(* IEC 61131-3 sources: daoli-st-library/DL_Process (part 4) *)

(* ---- FB_DL_MultiTankBlendSeq.st ---- *)
(*
  ============================================================
  组件名 : FB_DL_MultiTankBlendSeq
  分类   : DL_Process
  功能   : 多罐调和批次序列（A 进料 → B 进料 → 循环调和 → 取样 → 排料 → 完成），含超容、进料超时、收敛超时、取样超时、排料超时、人工中止、配方无效共七类故障锁存
  开源溯源 : internal-design（本轮无外部代码逐行引用）；参考语义 : 无外部参考
  复杂度 : C4
  版本   : 1.0.0
  ============================================================
*)

(*-----------------------------------------------------------------------------
 * 状态迁移表（ENUM 成员 → 出口；每成员均有可到达出口，零无界驻留相）：
 *   eIdle      → eFillA  : bStart 且 bRecipeValid 且组态闸通过 且 总量 ≤ rMaxVolume
 *   eIdle      ── 保持，直到 bStart（待机相以启动命令为唯一出口，属许可型驻留）
 *   eFillA     → eFillB  : rVolAct ≥ rVolA_sp（含 1E-6 容差）
 *   eFillA     → eFault  : tonFill.Q（码 1）｜bAbort 沿（码 5）｜rVolAct > rMaxVolume（码 4）｜bStart 撤除（无码回空闲）
 *   eFillB     → eCirculate : rVolAct ≥ (rVolA_sp + rVolB_sp) - 1E-6
 *   eFillB     → eFault  : tonFill.Q（码 1）｜bAbort 沿（码 5）｜超容（码 4）｜组态闸失效（码 6）
 *   eCirculate → eSample : 温度与浓度同时进带并持续 tCircStable（tonStable.Q）
 *   eCirculate → eFault  : tonCirc.Q（码 2）｜bAbort 沿（码 5）
 *   eSample    → eRelease : bSampleDone（外部取样完成电平）
 *   eSample    → eFault   : tonSample.Q（码 3）｜bAbort 沿（码 5）
 *   eRelease   → eDone    : bLevelLow（低液位信号，排料到位）
 *   eRelease   → eFault   : tonRelease.Q（码 7）｜bAbort 沿（码 5）
 *   eDone      → eIdle    : bStart 撤除（完成相以撤令为唯一出口，属人工确认型驻留）
 *   eFault     → eIdle    : bAbort 上升沿 或（bStart = FALSE 且 bAbort = FALSE）
 *   ELSE（非法枚举值，非任何成员）→ eFault（码 8）
 *
 * 故障码表（nFaultCode，0 = 无故障；非首码均附「现有输出不可观测」反证句，R90）：
 *   1 进料超时      : tFillTimeout 覆盖 eFillA + eFillB（进 eFillA 时计时器自然复位）。
 *   2 循环收敛超时  : 反证——eFault 相动作全撤后 bValveA/bValveB/bAgitator/bDischarge 全 FALSE、
 *                     eState 同为 eFault，复用码 1 会使「调和未收敛」与「进料过慢」在 HMI 上不可区分。
 *   3 取样超时      : 反证——取样相外部回执缺失，阀位与搅拌状态在故障撤除后与码 2 完全同形，
 *                     复用码 2 会把「外部取样单元不回报」误判为工艺收敛失败，运维方向相悖。
 *   4 超罐容        : 反证——超容判据在进料前即可成立（无阀位动作、无累计体积），
 *                     复用码 1 会把「配方总量超罐容」报成「进料慢」，掩盖配方错误。
 *   5 人工中止      : 反证——操作员主动撤令属安全审计事件，与任何超时码的因果主体不同，
 *                     合并后无法区分「设备不动」与「人按了停」。
 *   6 配方无效      : 反证——非法配方在进料前拦截，此时无累计体积、无阀位输出，
 *                     与超时类码位的时序签名互斥，必须独立成码以便前置拦截可被观测。
 *   7 排料超时      : 反证——排料相 bDischarge 独占且 bLevelLow 缺失，故障撤除后与码 1/2/3 的
 *                     观测量全同，复用码 1 会让运维去查进料阀而非排料阀。
 *   8 非法状态枚举  : 反证——非法枚举值为程序缺陷而非工艺事件，必须与现场工艺故障分离，
 *                     否则固件错误会被误排为设备故障。
 *
 * 依赖     : 仅 IEC 61131-3 标准库（TON / R_TRIG / ABS / LIMIT），零厂商私有库
 * 分工声明 : 循环泵输出不在本件接口（上层以 eState = eCirculate 派生泵命令）；
 *            温度/浓度闭环调节归温控件与浓度调节件；本件只做批次时序与保护，不做连续调节。
 * 归属     : E_DL_BlendState 归属本文件（全库唯一定义，R264；引用件只引用不重声明）。
 * 修订历史 : 2026-11-25  v1.0.0  首版（编码席 dlf-plc-coder，第二批 C4）
 *----------------------------------------------------------------------------*)

(*-----------------------------------------------------------------------------
 * 边界与红线自检：
 * ① 六个 TON 与一个 R_TRIG 全部在 CASE 外无条件周期调用（R7）；时间类 IN 均含 NOT .Q 自复位项
 *    与 NOT 故障锁存项（R188 / FB50-1③），CASE 内只读 .Q。
 * ② 出口命令（bValveA/bValveB/bAgitator/bDischarge/bSampleReq）在段 0 每拍预置 FALSE，
 *    CASE 内只置 TRUE —— eIdle 与 eFault 相零残留（上轮 MAJOR「故障后残留旧输出」型缺陷已封堵）。
 * ③ bDone 由相位派生（bDone := _eState = eDone），不是单拍脉冲，从结构上排除「同拍置位又撤销」（FB33-1）。
 * ④ 故障码 _nFault 一律锁存至 eFault 复位分支，故障相内不按当下输入重算（FB33-1③ / R152）。
 * ⑤ 除零防护：进度式除子 _rVolTotal 先过 > 1E-6 与 _bCfgOk 双检（R4）。
 * ⑥ 相内等待出口 ≥2（R98）：eSample = bSampleDone ｜ tonSample.Q ｜ bAbort 沿 ｜ bStart 撤除；
 *    eRelease = bLevelLow ｜ tonRelease.Q ｜ bAbort 沿 ｜ bStart 撤除。
 * ⑦ 组态域闸：参与任何判据换算的 10 个浮点入参全部显式枚举（含 rMaxVolume），NaN 用自反比较、
 *    Inf 用差值自减双判（R151 / R79），非有限不入保持槽。
 * ⑧ 零全局耦合：无 GVL / VAR_EXTERNAL / %I / %Q（R1 / R2）。
 * ⑨ 相位写入点共三处且互斥：段 3（bAbort 沿只置锁存，不写相位）、段 4 CASE、段 6 迁移闸。
 *----------------------------------------------------------------------------*)

TYPE E_DL_BlendState :
(
    eIdle      := 0, // 空闲：全部阀位关闭，等启动与配方有效 idle: all valves closed, waiting for start and a valid recipe
    eFillA     := 1, // A 罐进料相：开 A 阀累计至 rVolA_sp fill A: A valve open until rVolA_sp is reached
    eFillB     := 2, // B 罐进料相：开 B 阀累计至 A+B 总量 fill B: B valve open until the A+B total is reached
    eCirculate := 3, // 循环调和相：搅拌运行，温度与浓度双判进带 circulate: agitation with temperature and concentration both inside band
    eSample    := 4, // 取样相：置取样请求等外部完成 sample: sample request raised, waiting for the external completion
    eRelease   := 5, // 排料相：开排料阀至低液位 release: discharge valve open until the low level signal
    eFault     := 6, // 故障锁存相：全部阀位撤除，只由复位出口迁出 fault: all valves withdrawn, left only by the reset outlet
    eDone      := 7  // 批次完成相：bStart 撤除后回空闲 done: returns to idle when bStart is withdrawn
);
END_TYPE

FUNCTION_BLOCK FB_DL_MultiTankBlendSeq
VAR_INPUT
    bStart          : BOOL := FALSE;          // 启动/运行许可（电平）：撤除即安全停机回空闲 [bool] start and run permissive, a dropped level stops safely
    bAbort          : BOOL := FALSE;          // 人工中止（上升沿）：置故障码 5 并锁存 [bool] manual abort rising edge, latches fault code 5
    bRecipeValid    : BOOL := FALSE;          // 配方有效回执：FALSE 时禁止启动并置码 6 [bool] recipe valid receipt, FALSE blocks the start with code 6
    rVolA_sp        : REAL := 0.0;            // A 组分配方体积设定 [m3] recipe volume setpoint of component A [m3]
    rVolB_sp        : REAL := 0.0;            // B 组分配方体积设定 [m3] recipe volume setpoint of component B [m3]
    rVolAct         : REAL := 0.0;            // 当前累计进料量（A+B 合计）[m3] accumulated feed volume of A plus B [m3]
    rTempAct        : REAL := 0.0;            // 混合物实测温度 [degC] measured blend temperature [degC]
    rTempSp         : REAL := 0.0;            // 调和温度设定 [degC] blend temperature setpoint [degC]
    rTempBand       : REAL := 0.0;            // 温度进带允许偏差，域 > 1E-6 [K] temperature band tolerance, domain > 1E-6 [K]
    rConcAct        : REAL := 0.0;            // 混合物实测浓度 [%] measured blend concentration [%]
    rConcSp         : REAL := 0.0;            // 调和浓度设定 [%] blend concentration setpoint [%]
    rConcBand       : REAL := 0.0;            // 浓度进带允许偏差，域 > 1E-6 [%] concentration band tolerance, domain > 1E-6 [%]
    tFillTimeout    : TIME := T#10M;          // 进料总超时窗，覆盖 eFillA + eFillB [s] total feed timeout covering fill A and fill B [s]
    tCircTimeout    : TIME := T#30M;          // 循环调和相超时窗 [s] circulation phase timeout window [s]
    tSampleTimeout  : TIME := T#5M;           // 取样相等待外部回执超时窗 [s] sample phase external receipt timeout [s]
    rMaxVolume      : REAL := 10.0;           // 罐体最大有效容积，域 > 0 [m3] tank maximum usable volume, domain > 0 [m3]
    bSampleDone     : BOOL := FALSE;          // 外部取样完成回执（电平）[bool] external sampling done receipt level
    bLevelLow       : BOOL := FALSE;          // 排料低液位信号（排料到位）[bool] discharge low level signal
    tCircStable     : TIME := T#15S;          // 温度与浓度同时在带内的持续确认窗 [s] continuous in-band confirmation window [s]
    tReleaseTimeout : TIME := T#15M;          // 排料相超时窗（低液位不到的兜底）[s] release phase timeout fallback [s]
END_VAR
VAR_OUTPUT
    bValveA      : BOOL;                      // A 组分进料阀命令（段 0 预置，CASE 只置位）[bool] component A feed valve command
    bValveB      : BOOL;                      // B 组分进料阀命令（段 0 预置，CASE 只置位）[bool] component B feed valve command
    bAgitator    : BOOL;                      // 搅拌器命令（循环相与取样相保持开）[bool] agitator command, held in circulation and sampling
    bDischarge   : BOOL;                      // 排料阀命令（仅排料相）[bool] discharge valve command, release phase only
    bSampleReq   : BOOL;                      // 取样请求（仅取样相，电平保持）[bool] sample request, level held in the sample phase
    eState       : E_DL_BlendState;           // 相位出口（段 7 单点映射）[-] phase outlet mapped once in section 7
    bDone        : BOOL;                      // 批次完成（由相位派生，非单拍脉冲）[bool] batch done, derived from the phase as a level
    nFaultCode   : INT;                       // 故障码 0 无 1 进料超时 2 收敛超时 3 取样超时 4 超容 5 人工中止 6 配方无效 7 排料超时 8 非法状态 [码] fault code
    rProgressPct : REAL;                      // 进料完成度 0..100（其后各相恒 100）[%] feed completion percentage, constant 100 in later phases [%]
    bError       : BOOL;                      // 故障锁存标志（取锁存位，R45 配对出口）[bool] fault latch flag used as the paired outlet
END_VAR
VAR
    _eState       : E_DL_BlendState := E_DL_BlendState.eIdle;   // 内部相位（CASE 唯一比较目标）[-] internal phase compared by the CASE
    _bFaultLatch  : BOOL := FALSE;                              // 故障锁存位（仅复位出口清除）[bool] fault latch, cleared only by the reset outlet
    _nFault       : INT := 0;                                   // 锁存故障码（故障期回放，不按当下输入重算）[码] latched fault code replayed during the fault phase
    _bCfgOk       : BOOL := FALSE;                              // 组态与入参域闸通过标志 [bool] configuration and input domain gate flag
    _bRunActive   : BOOL := FALSE;                              // 运行相关相标志（进料到排料）[bool] running phase flag from fill to release
    _bInBand      : BOOL := FALSE;                               // 温度与浓度同时进带标志 [bool] both temperature and concentration inside band
    _bValveA      : BOOL := FALSE;                              // 内部 A 阀命令状态 [bool] internal A valve command state
    _bValveB      : BOOL := FALSE;                              // 内部 B 阀命令状态 [bool] internal B valve command state
    _bAgitator    : BOOL := FALSE;                              // 内部搅拌命令状态 [bool] internal agitator command state
    _bDischarge   : BOOL := FALSE;                              // 内部排料阀命令状态 [bool] internal discharge valve command state
    _bSampleReq   : BOOL := FALSE;                              // 内部取样请求状态 [bool] internal sample request state
    _rVolTotal    : REAL := 0.0;                                // 配方总量 = A + B [m3] recipe total volume of A plus B [m3]
    _rProg        : REAL := 0.0;                                // 进料完成度中间量 [%] feed completion intermediate value [%]
    rtAbort       : R_TRIG;                                     // bAbort 上升沿实例（段 2 无条件调用）[bool] abort rising edge instance
    tonFill       : TON;                                        // 进料总超时计时（覆盖两进料相，段 2 无条件调用）[s] total feed timeout covering both fill phases
    tonCirc       : TON;                                        // 循环调和相超时计时（段 2 无条件调用）[s] circulation timeout
    tonStable     : TON;                                        // 双判进带持续确认计时（段 2 无条件调用）[s] in-band persistence timer
    tonSample     : TON;                                        // 取样相等待回执超时计时（段 2 无条件调用）[s] sample receipt timeout
    tonRelease    : TON;                                        // 排料相超时计时（段 2 无条件调用）[s] release timeout
END_VAR
VAR CONSTANT
    DL_BLD_ZERO     : REAL := 0.0;        // 浮点零基准 [m3] float zero base
    DL_BLD_ONE      : REAL := 1.0;        // 浮点一基准 [%] float one base
    DL_BLD_HUNDRED  : REAL := 100.0;      // 百分比满量程 [%] percent full scale
    DL_BLD_EPS      : REAL := 1.0E-6;     // 体积与宽容差基准 [m3] volume and band tolerance base
    DL_BLD_T_MIN    : TIME := T#100MS;    // 时间参数下限 [s] lower bound of the time parameters
    DL_BLD_T_MAX    : TIME := T#4H;       // 时间参数上限 [s] upper bound of the time parameters
END_VAR

(* —— 段 0：出口命令预置与派生量计算（CASE 内只置 TRUE，杜绝故障相残留） —— *)
_bValveA    := FALSE;                                               // A 阀命令每拍先撤 [bool] A valve withdrawn first each scan
_bValveB    := FALSE;                                               // B 阀命令每拍先撤 [bool] B valve withdrawn first each scan
_bAgitator  := FALSE;                                               // 搅拌命令每拍先撤 [bool] agitator withdrawn first each scan
_bDischarge := FALSE;                                               // 排料阀命令每拍先撤 [bool] discharge withdrawn first each scan
_bSampleReq := FALSE;                                               // 取样请求每拍先撤 [bool] sample request withdrawn first each scan
_rProg      := DL_BLD_ZERO;                                         // 进度中间量每拍清零 [%] progress intermediate cleared each scan
_rVolTotal  := rVolA_sp + rVolB_sp;                                 // 配方总量求和 [m3] recipe total volume
_bRunActive := (_eState = E_DL_BlendState.eFillA) OR (_eState = E_DL_BlendState.eFillB)
               OR (_eState = E_DL_BlendState.eCirculate) OR (_eState = E_DL_BlendState.eSample)
               OR (_eState = E_DL_BlendState.eRelease);             // 运行相关相标志（用状态量，R99）[bool] running phase flag from the state
_bInBand    := FALSE;                                               // 进带标志复位 [bool] in-band flag reset
IF (rTempBand > DL_BLD_ZERO) AND (rConcBand > DL_BLD_ZERO) THEN
    IF (ABS(rTempAct - rTempSp) <= rTempBand) AND (ABS(rConcAct - rConcSp) <= rConcBand) THEN
        _bInBand := TRUE;                                           // 双判同时进带 [bool] both criteria inside band
    END_IF
END_IF

(* —— 段 1：组态域闸与容量保护（十个浮点入参全枚举，非有限双判 R151 / R79） —— *)
_bCfgOk := TRUE;                                                    // 组态闸标志初值 [bool] configuration flag initial value
IF (rVolA_sp <> rVolA_sp) OR ((rVolA_sp - rVolA_sp) <> DL_BLD_ZERO)
   OR (rVolB_sp <> rVolB_sp) OR ((rVolB_sp - rVolB_sp) <> DL_BLD_ZERO)
   OR (rVolAct <> rVolAct) OR ((rVolAct - rVolAct) <> DL_BLD_ZERO)
   OR (rMaxVolume <> rMaxVolume) OR ((rMaxVolume - rMaxVolume) <> DL_BLD_ZERO)
   OR (rTempAct <> rTempAct) OR ((rTempAct - rTempAct) <> DL_BLD_ZERO)
   OR (rTempSp <> rTempSp) OR ((rTempSp - rTempSp) <> DL_BLD_ZERO)
   OR (rTempBand <> rTempBand) OR ((rTempBand - rTempBand) <> DL_BLD_ZERO)
   OR (rConcAct <> rConcAct) OR ((rConcAct - rConcAct) <> DL_BLD_ZERO)
   OR (rConcSp <> rConcSp) OR ((rConcSp - rConcSp) <> DL_BLD_ZERO)
   OR (rConcBand <> rConcBand) OR ((rConcBand - rConcBand) <> DL_BLD_ZERO) THEN
    _bCfgOk := FALSE;                                               // 非有限入参：拒收（NaN 自反 + Inf 差值自减）[bool] non finite input rejected
END_IF
IF _bCfgOk THEN
    IF (rVolA_sp < DL_BLD_ZERO) OR (rVolB_sp < DL_BLD_ZERO) OR (rMaxVolume <= DL_BLD_ZERO) THEN
        _bCfgOk := FALSE;                                           // 负体积或非正罐容 [bool] negative volume or non positive capacity
    ELSIF (_rVolTotal <= DL_BLD_ZERO) THEN
        _bCfgOk := FALSE;                                           // 配方总量为零 [bool] zero recipe total volume
    ELSIF (rTempBand < DL_BLD_EPS) OR (rConcBand < DL_BLD_EPS) THEN
        _bCfgOk := FALSE;                                           // 容差带为零或负 [bool] zero or negative tolerance band
    ELSIF (tFillTimeout < DL_BLD_T_MIN) OR (tFillTimeout > DL_BLD_T_MAX) THEN
        _bCfgOk := FALSE;                                           // 进料超时越域 [bool] feed timeout out of domain
    ELSIF (tCircTimeout < DL_BLD_T_MIN) OR (tCircTimeout > DL_BLD_T_MAX) THEN
        _bCfgOk := FALSE;                                           // 循环超时越域 [bool] circulation timeout out of domain
    ELSIF (tSampleTimeout < DL_BLD_T_MIN) OR (tSampleTimeout > DL_BLD_T_MAX) THEN
        _bCfgOk := FALSE;                                           // 取样超时越域 [bool] sample timeout out of domain
    ELSIF (tCircStable < DL_BLD_T_MIN) OR (tCircStable > DL_BLD_T_MAX) THEN
        _bCfgOk := FALSE;                                           // 进带确认窗越域 [bool] in-band window out of domain
    ELSIF (tReleaseTimeout < DL_BLD_T_MIN) OR (tReleaseTimeout > DL_BLD_T_MAX) THEN
        _bCfgOk := FALSE;                                           // 排料超时越域 [bool] release timeout out of domain
    ELSIF NOT bRecipeValid THEN
        _bCfgOk := FALSE;                                           // 配方无效回执为假 [bool] recipe valid receipt is false
    END_IF
END_IF
IF (NOT _bCfgOk) AND (NOT _bFaultLatch) AND (bStart OR _bRunActive) THEN
    _nFault      := 6;                                              // 故障级：配方无效 / 参数非法 [码] fault: invalid recipe or parameter
    _bFaultLatch := TRUE;                                           // 置故障锁存 [bool] latch the fault
    bError       := TRUE;                                           // R45 配对：故障标志同拍置位 [bool] paired error flag
END_IF
IF (NOT _bFaultLatch) AND (bStart OR _bRunActive) THEN
    IF _rVolTotal > rMaxVolume THEN
        _nFault      := 4;                                          // 故障级：配方总量超罐容 [码] fault: recipe total exceeds tank volume
        _bFaultLatch := TRUE;                                       // 置故障锁存 [bool] latch the fault
        bError       := TRUE;                                       // R45 配对：故障标志同拍置位 [bool] paired error flag
    END_IF
END_IF

(* —— 段 2：边沿与定时器（CASE 外无条件周期调用，R7；IN 含 NOT .Q 自复位与 NOT 锁存，R188） —— *)
rtAbort(CLK := bAbort);                                             // bAbort 边沿无条件刷新 [bool] abort edge refreshed unconditionally
tonFill(IN := ((_eState = E_DL_BlendState.eFillA) OR (_eState = E_DL_BlendState.eFillB))
              AND (NOT tonFill.Q) AND (NOT _bFaultLatch),
        PT := tFillTimeout);                                        // 进料总超时（跨两相累计，进相自然复位）[s] total feed timeout across both phases
tonCirc(IN := (_eState = E_DL_BlendState.eCirculate) AND (NOT tonCirc.Q) AND (NOT _bFaultLatch),
        PT := tCircTimeout);                                        // 循环调和超时 [s] circulation timeout
tonStable(IN := (_eState = E_DL_BlendState.eCirculate) AND _bInBand AND (NOT tonStable.Q)
               AND (NOT _bFaultLatch),
          PT := tCircStable);                                       // 双判进带持续确认 [s] in-band persistence confirmation
tonSample(IN := (_eState = E_DL_BlendState.eSample) AND (NOT tonSample.Q) AND (NOT _bFaultLatch),
          PT := tSampleTimeout);                                    // 取样回执超时 [s] sample receipt timeout
tonRelease(IN := (_eState = E_DL_BlendState.eRelease) AND (NOT tonRelease.Q) AND (NOT _bFaultLatch),
           PT := tReleaseTimeout);                                  // 排料超时 [s] release timeout

(* —— 段 3：人工中止优先消化（置锁存不写相位，迁相由段 6 统一执行，R21 / R275） —— *)
IF rtAbort.Q AND (NOT _bFaultLatch) THEN
    _nFault      := 5;                                              // 故障级：人工中止 [码] fault: manual abort
    _bFaultLatch := TRUE;                                           // 置故障锁存 [bool] latch the fault
    bError       := TRUE;                                           // R45 配对：故障标志同拍置位 [bool] paired error flag
END_IF

(* —— 段 4：主状态机（相位写入点之二；每成员独立标签，ELSE 只兜非法值） —— *)
CASE _eState OF
E_DL_BlendState.eIdle :                                             // 空闲相：全部阀位已撤，等启动与配方许可
    IF bStart AND _bCfgOk AND (NOT bAbort) AND (NOT _bFaultLatch) THEN
        _eState := E_DL_BlendState.eFillA;                          // 迁移：进入 A 进料相（次拍开阀）[phase] move to fill A
    END_IF

E_DL_BlendState.eFillA :                                            // A 进料相：开 A 阀
    _bValveA := TRUE;                                               // 开 A 组分进料阀 [bool] open the component A feed valve
    IF rVolAct >= (rVolA_sp - DL_BLD_EPS) THEN
        _eState := E_DL_BlendState.eFillB;                          // 迁移：A 组分量已到位 [phase] component A volume reached
    ELSIF rVolAct > rMaxVolume THEN
        _nFault      := 4;                                          // 故障级：累计体积超罐容 [码] fault: accumulated volume over capacity
        _bFaultLatch := TRUE;                                       // 置故障锁存 [bool] latch the fault
        bError       := TRUE;                                       // R45 配对：故障标志同拍置位 [bool] paired error flag
    END_IF

E_DL_BlendState.eFillB :                                            // B 进料相：开 B 阀至总量
    _bValveB := TRUE;                                               // 开 B 组分进料阀 [bool] open the component B feed valve
    IF rVolAct >= (_rVolTotal - DL_BLD_EPS) THEN
        _eState := E_DL_BlendState.eCirculate;                      // 迁移：总量到位进入循环调和 [phase] total volume reached, start circulation
    ELSIF rVolAct > rMaxVolume THEN
        _nFault      := 4;                                          // 故障级：累计体积超罐容 [码] fault: accumulated volume over capacity
        _bFaultLatch := TRUE;                                       // 置故障锁存 [bool] latch the fault
        bError       := TRUE;                                       // R45 配对：故障标志同拍置位 [bool] paired error flag
    END_IF

E_DL_BlendState.eCirculate :                                        // 循环调和相：搅拌运行，温度与浓度双判
    _bAgitator := TRUE;                                             // 搅拌保持开（保证均质）[bool] agitator held on for homogeneity
    IF tonStable.Q THEN
        _eState := E_DL_BlendState.eSample;                         // 迁移：双判进带持续满足 [phase] both criteria held inside band
    END_IF

E_DL_BlendState.eSample :                                           // 取样相：请求外部取样并等待回执
    _bAgitator  := TRUE;                                            // 取样期间保持搅拌（样品代表性）[bool] agitator held during sampling
    _bSampleReq := TRUE;                                            // 置取样请求（电平保持）[bool] sample request level held
    IF bSampleDone THEN
        _eState := E_DL_BlendState.eRelease;                        // 迁移（出口 1）：外部取样完成 [phase] external sampling completed
    END_IF

E_DL_BlendState.eRelease :                                          // 排料相：开排料阀至低液位
    _bDischarge := TRUE;                                            // 开排料阀（搅拌停，避免抽空涡流）[bool] open the discharge valve
    IF bLevelLow THEN
        _eState := E_DL_BlendState.eDone;                           // 迁移（出口 1）：低液位到位 [phase] low level reached
    END_IF

E_DL_BlendState.eDone :                                             // 完成相：bDone 由相位派生，等撤令
    IF NOT bStart THEN
        _eState := E_DL_BlendState.eIdle;                           // 迁移：撤除启动命令回空闲 [phase] start withdrawn, back to idle
    END_IF

E_DL_BlendState.eFault :                                            // 故障锁存相：阀位已由段 6 全撤
    IF rtAbort.Q OR ((NOT bStart) AND (NOT bAbort)) THEN
        _bFaultLatch := FALSE;                                      // 复位出口：清故障锁存 [bool] clear the fault latch
        _nFault      := 0;                                          // 复位出口：清故障码 [码] clear the fault code
        _eState      := E_DL_BlendState.eIdle;                      // 复位出口：迁回空闲 [phase] back to idle
    END_IF

ELSE                                                                // 非法枚举值兜底（R6 / FB32-5）
    IF NOT _bFaultLatch THEN
        _nFault      := 8;                                          // 故障级：非法状态枚举值 [码] fault: illegal state enum value
        _bFaultLatch := TRUE;                                       // 置故障锁存 [bool] latch the fault
        bError       := TRUE;                                       // R45 配对：故障标志同拍置位 [bool] paired error flag
    END_IF
    _eState := E_DL_BlendState.eFault;                              // 非法值一律落安全相 [phase] illegal value falls into the safe phase
END_CASE

(* —— 段 5：超时看门狗锁存（本拍合法事件优先于超时：状态已迁出则该相看门狗不生效，R275） —— *)
IF tonFill.Q AND (NOT _bFaultLatch)
   AND ((_eState = E_DL_BlendState.eFillA) OR (_eState = E_DL_BlendState.eFillB)) THEN
    _nFault      := 1;                                              // 故障级：进料超时 [码] fault: feed timeout
    _bFaultLatch := TRUE;                                           // 置故障锁存 [bool] latch the fault
    bError       := TRUE;                                           // R45 配对：故障标志同拍置位 [bool] paired error flag
END_IF
IF tonCirc.Q AND (NOT _bFaultLatch) AND (_eState = E_DL_BlendState.eCirculate) THEN
    _nFault      := 2;                                              // 故障级：循环收敛超时 [码] fault: circulation convergence timeout
    _bFaultLatch := TRUE;                                           // 置故障锁存 [bool] latch the fault
    bError       := TRUE;                                           // R45 配对：故障标志同拍置位 [bool] paired error flag
END_IF
IF tonSample.Q AND (NOT _bFaultLatch) AND (_eState = E_DL_BlendState.eSample) THEN
    _nFault      := 3;                                              // 故障级：取样超时 [码] fault: sampling timeout
    _bFaultLatch := TRUE;                                           // 置故障锁存 [bool] latch the fault
    bError       := TRUE;                                           // R45 配对：故障标志同拍置位 [bool] paired error flag
END_IF
IF tonRelease.Q AND (NOT _bFaultLatch) AND (_eState = E_DL_BlendState.eRelease) THEN
    _nFault      := 7;                                              // 故障级：排料超时 [码] fault: release timeout
    _bFaultLatch := TRUE;                                           // 置故障锁存 [bool] latch the fault
    bError       := TRUE;                                           // R45 配对：故障标志同拍置位 [bool] paired error flag
END_IF

(* —— 段 6：段尾故障迁移闸 + 撤令安全停机 + 故障/空闲相动作全撤（FB50-1④ / R191 显式声明） —— *)
IF _bFaultLatch AND (_eState <> E_DL_BlendState.eFault) THEN
    _eState := E_DL_BlendState.eFault;                              // 锁存即迁相（锁存与迁相分离，R21）[phase] a latch forces the fault phase
END_IF
IF (NOT bStart) AND _bRunActive AND (NOT _bFaultLatch) THEN
    (* 撤令语义（R191 二选一，本件选「降级为安全值 + 回空闲，不置故障码」）：阀位全撤、相位回空闲 *)
    _eState := E_DL_BlendState.eIdle;                               // 撤令即安全停机回空闲 [phase] withdrawn start stops safely into idle
END_IF
IF (_eState = E_DL_BlendState.eFault) OR (_eState = E_DL_BlendState.eIdle) THEN
    _bValveA    := FALSE;                                           // 空闲/故障：A 阀全撤 [bool] A valve withdrawn in idle and fault
    _bValveB    := FALSE;                                           // 空闲/故障：B 阀全撤 [bool] B valve withdrawn in idle and fault
    _bAgitator  := FALSE;                                           // 空闲/故障：搅拌全撤 [bool] agitator withdrawn in idle and fault
    _bDischarge := FALSE;                                           // 空闲/故障：排料阀全撤 [bool] discharge withdrawn in idle and fault
    _bSampleReq := FALSE;                                           // 空闲/故障：取样请求撤除 [bool] sample request withdrawn in idle and fault
END_IF

(* —— 段 7：统一出口（相位映射 + 进度换算 + 锁存码回放；单一写入点） —— *)
IF ((_eState = E_DL_BlendState.eFillA) OR (_eState = E_DL_BlendState.eFillB)) AND _bCfgOk THEN
    IF _rVolTotal > DL_BLD_EPS THEN
        _rProg := LIMIT(DL_BLD_ZERO, (rVolAct * DL_BLD_HUNDRED) / _rVolTotal, DL_BLD_HUNDRED); // 进料完成度（除子已双检，R4）[%] feed completion
    END_IF
ELSIF (_eState = E_DL_BlendState.eCirculate) OR (_eState = E_DL_BlendState.eSample)
   OR (_eState = E_DL_BlendState.eRelease) OR (_eState = E_DL_BlendState.eDone) THEN
    _rProg := DL_BLD_HUNDRED;                                       // 进料已完成，其后各相进度满量程 [%] feed finished, later phases at full scale
END_IF
bValveA      := _bValveA;                                           // A 阀命令出口 [bool] A valve command outlet
bValveB      := _bValveB;                                           // B 阀命令出口 [bool] B valve command outlet
bAgitator    := _bAgitator;                                         // 搅拌命令出口 [bool] agitator command outlet
bDischarge   := _bDischarge;                                        // 排料阀命令出口 [bool] discharge command outlet
bSampleReq   := _bSampleReq;                                        // 取样请求出口 [bool] sample request outlet
eState       := _eState;                                            // 相位出口 [phase] phase outlet
bDone        := (_eState = E_DL_BlendState.eDone);                  // 完成位由相位派生（非单拍脉冲）[bool] done derived from the phase
nFaultCode   := _nFault;                                            // 故障码出口（锁存回放）[码] fault code outlet replayed from the latch
rProgressPct := _rProg;                                             // 进度出口 [%] progress outlet
bError       := _bFaultLatch;                                       // 故障标志取锁存位 [bool] fault flag from the latch
END_FUNCTION_BLOCK

(* ---- FB_DL_OcvTempNormalize.st ---- *)
(*==============================================================================
 * 组件名称 (Component)  : FB_DL_OcvTempNormalize
 * 所属子库 (Sublibrary) : DL_Process
 * 当前版本 (Version)    : 1.0.0
 * 兼容性   (Platform)   : CODESYS 3.5+ / TwinCAT 3 / 汇川 InoProShop / 施耐德 Machine Expert
 *                         仅依赖 Standard.library（R_TRIG），零厂商私有库
 * 功能描述 (Function)   : OCV（开路电压）测试温度归一判据。
 *                         把实测 OCV 按温度系数线性归一到基准温度，再对归一值做合格带判定与三档分级。
 *                         归一式（一阶线性，符号约定写死）：
 *                           OCV_norm = OCV_meas + k · (T_meas − T_ref)
 *                           其中 k 为温度系数 [mV/°C]，正值表示"温度升高时实测 OCV 升高"，
 *                           故归一化需回减 k·ΔT；k 为负（低温型电芯）同样成立，不做符号假设。
 *                         **语义复用（非实例复用）**：按 R47 批次"批内零 .st 文件级依赖"纪律，
 *                         不实例化 FC_DL_TempUnitConvert，而复用其已固化的三条换算语义——
 *                         ① 华氏 → 摄氏用 (F−32)·5/9；② 开尔文 → 摄氏用 K−273.15；
 *                         ③ 未知单位一律拒绝换算并置故障级（不猜默认单位）。
 *                         验收向量：
 *                           ① OCV=3850 mV, T=35 °C, k=+0.5 mV/°C, Tref=25 °C
 *                              → 归一 = 3850 + 0.5×(35−25) = 3855 mV
 *                           ② OCV=3850 mV, T=25 °C → 归一 = 3850 mV（ΔT=0，归一不改变量值）
 *                           ③ 带 [3800, 3900] mV，归一 3855 → eInBand；3901 → eHigh；3799 → eLow
 *                           ④ k=0 → 拒归一（除零语义的乘法侧等价：k=0 时归一退化，判据失真）
 * 接口     (Interface)  : 入 bEnable 使能（FALSE 冻结判据且不宣称）、fOcvMeasMv 实测 OCV、fTempMeas
 *                         实测温度、iTempUnit 温度单位、fTempCoeff 温度系数、fTempRefC 基准温度、
 *                         fBandLowMv / fBandHighMv 合格带上下限、fNormClampMv 归一值钳位、
 *                         bReset 故障复位沿；
 *                         出 fOcvNormMv 归一后 OCV、bInBand 合格、eGrade 三档分级、
 *                         bValid 结果有效、eState 相、eCause 成因、bError 故障标志。
 * 边界     (Boundary)   : ① **属主边界（写死）：本件只做"归一 + 判带"，不判电芯合格结论
 *                         （那是分选件的最终裁决），不做 OCV 采样时序、不驱动测试仪**；
 *                         ② **温度系数零闸**：k 为 0（或非有限）→ 归一退化，锁存 eCoeffZero，
 *                         判据整体停用（静默失效比报错危险，R179）；
 *                         ③ **合格带倒置闸**：fBandLow ≥ fBandHigh → 锁存 eCfgIllegal；
 *                         ④ **钳位**：归一值超 ±fNormClampMv 时钳位并置 bClamped（脚非法时回退
 *                         VAR CONSTANT，R127 兜底与判定量解耦）；
 *                         ⑤ **非有限样本**：OCV / 温度任一非有限 → 当拍不判、bValid=FALSE、
 *                         不锁存（可恢复性瞬时异常，与组态类锁存分轨，R228B）；
 *                         ⑥ 浮点比较一律差值容差判等（本件判带用 ABS 差 < fEps）；
 *                         ⑦ eFault 可迁出：bReset 上升沿 → eIdle，解除式恒可达（外部引脚门控）；
 *                         ⑧ 零全局耦合、零物理地址。
 * 分工声明 (Scope)      : 本件只管"温度归一与合格带判定"。不接管：温补分档迟滞
 *                         （属 FB_DL_TempCompClassify）、电芯分选结论（属分选件）、
 *                         温度采集与滤波（属模拟量通道件）。
 * 来源标签 (Source Tag) : ROADMAP 空勾真缺口 P1（OCV 温度归一，自研 clean-room）
 * 码表     (Codes)      : 本件不占用任何全局数字码位（零码位范式 R297）；诊断由 BOOL + ENUM 出口承担。
 * 红线自检 (Redline)    : R1 ✓ 零 GVL/VAR_EXTERNAL ｜ R2 ✓ 零 %I/%Q/%M ｜ R3 ✓ 纯 IEC 61131-3
 *                         R4 ✓ 零闸 + 倒置闸 + 钳位 + 非有限闸 + 容差判等 ｜ R5 ✓ 声明逐行同行双语注释
 *                         R6 ✓ ENUM+CASE 含 ELSE 兜底 ｜ R7 ✓ R_TRIG 段 0 无条件刷新（本件无 TON）
 * 修订历史 (Revision)   : 2026-11-19  v1.0.0  R47 首版（批次 1 · 序号 5）
 *==============================================================================*)

TYPE E_DL_OtnUnit :
(
    eCelsius    := 0,   // 摄氏（本件内部基准单位） / Celsius, the internal base unit
    eFahrenheit := 1,   // 华氏 / Fahrenheit
    eKelvin     := 2,   // 开尔文 / Kelvin
    eUnknown    := 3    // 未知单位（拒换算，故障级） / Unknown unit, conversion refused
);
END_TYPE

TYPE E_DL_OtnGrade :
(
    eNoGrade := 0,   // 未分级（无效或未使能） / Ungraded, invalid or disabled
    eLow     := 1,   // 低于合格带（归一值偏低） / Below the accept band
    eInBand  := 2,   // 落合格带内 / Inside the accept band
    eHigh    := 3    // 高于合格带（归一值偏高） / Above the accept band
);
END_TYPE

TYPE E_DL_OtnState :
(
    eIdle  := 0,    // 待机相（未使能） / Idle, disabled
    eRun   := 10,   // 判据相（归一与判带） / Running, normalise and classify
    eFault := 90    // 故障相（等复位） / Fault, awaiting reset
);
END_TYPE

TYPE E_DL_OtnCause :
(
    eNone      := 0,   // 无异常 / No anomaly
    eCfgIllegal:= 1,   // 组态非法（合格带倒置/钳位限非正） / Illegal configuration
    eCoeffZero := 2,   // 温度系数为零（归一退化，拒判） / Zero temperature coefficient
    eUnitBad   := 3,   // 温度单位未知（拒换算） / Unknown temperature unit
    ePhaseBad  := 4    // 非法相位兜底 / Illegal phase fallback
);
END_TYPE

FUNCTION_BLOCK FB_DL_OcvTempNormalize
VAR_INPUT
    bEnable      : BOOL := FALSE;        // 使能（FALSE 冻结判据且不宣称） [-] / Enable, freezes the judgement when FALSE
    fOcvMeasMv   : LREAL := 0.0;         // 实测 OCV [mV] / Measured open-circuit voltage [mV]
    fTempMeas    : LREAL := 25.0;        // 实测温度（按 iTempUnit 解释） [°C/°F/K] / Measured temperature in the declared unit
    iTempUnit    : E_DL_OtnUnit := E_DL_OtnUnit.eCelsius;   // 温度单位 [-] / Temperature unit
    fTempCoeff   : LREAL := 0.5;         // 温度系数 k，域 ≠ 0 [mV/°C] / Temperature coefficient, non-zero
    fTempRefC    : LREAL := 25.0;        // 基准温度（摄氏） [°C] / Reference temperature in Celsius
    fBandLowMv   : LREAL := 3800.0;      // 合格带下限 [mV] / Accept band lower limit [mV]
    fBandHighMv  : LREAL := 3900.0;      // 合格带上限，域 > 下限 [mV] / Accept band upper limit [mV]
    fNormClampMv : LREAL := 30000.0;     // 归一值绝对钳位，域 > 0 [mV] / Absolute clamp of the normalised value
    bReset       : BOOL := FALSE;        // 故障复位沿 [-] / Fault reset edge
END_VAR
VAR_OUTPUT
    fOcvNormMv : LREAL := 0.0;                       // 归一到基准温度后的 OCV [mV] / OCV normalised to the reference temperature
    bInBand    : BOOL := FALSE;                      // 归一值落合格带内 [-] / Normalised value inside the accept band
    eGrade     : E_DL_OtnGrade := E_DL_OtnGrade.eNoGrade;   // 三档分级出口 [-] / Three-way grade outlet
    bValid     : BOOL := FALSE;                      // 结果有效（样本有限且已归一） [-] / Result valid
    bClamped   : BOOL := FALSE;                      // 归一值被钳位 [-] / Normalised value clamped
    eState     : E_DL_OtnState := E_DL_OtnState.eIdle;      // 相出口 [-] / Phase outlet
    eCause     : E_DL_OtnCause := E_DL_OtnCause.eNone;      // 成因出口（R190 归因唯一） [-] / Cause outlet
    bError     : BOOL := FALSE;                      // 故障标志 [-] / Error flag
END_VAR
VAR
    _eState  : E_DL_OtnState := E_DL_OtnState.eIdle;        // 内部相（CASE 唯一写入目标） / Internal phase
    _eCause  : E_DL_OtnCause := E_DL_OtnCause.eNone;        // 成因锁存量 / Latched cause
    _bFault  : BOOL := FALSE;                               // 故障锁存位 / Latched fault bit
    _fTempC  : LREAL := 0.0;                                // 换算后的摄氏温度 [°C] / Temperature converted to Celsius
    _fNorm   : LREAL := 0.0;                                // 归一计算工作值 [mV] / Normalisation working value
    _fLim    : LREAL := 0.0;                                // 生效钳位限（脚非法回退常量，R127） [mV] / Effective clamp limit
    _bXFin   : BOOL := FALSE;                               // 样本有限性判定中间量 [-] / Sample finiteness working flag
    _bBandOk : BOOL := FALSE;                               // 合格带域闸结论 [-] / Accept-band domain gate result
    rtReset  : R_TRIG;                                      // 复位沿实例，段 0 无条件调用 / Reset edge instance
END_VAR
VAR CONSTANT
    DL_OTN_CLAMP_DEF : LREAL := 30000.0;    // 钳位限回退默认值（与脚默认同源） [mV] / Default clamp limit
    DL_OTN_K2C       : LREAL := 273.15;     // 开尔文转摄氏偏移量 [°C] / Kelvin-to-Celsius offset
    DL_OTN_F_SCALE   : LREAL := 5.0 / 9.0;  // 华氏温差换算比例（5/9，常量预算不除零） [-] / Fahrenheit delta ratio
    DL_OTN_F_OFFS    : LREAL := 32.0;       // 华氏冰点偏移 [°F] / Fahrenheit ice-point offset
    DL_OTN_EPS       : LREAL := 1.0E-6;     // 浮点判等容差（仅用于"贴带边"判定） [mV] / Equality tolerance
END_VAR

(* —— 段 0：两枚沿实例无条件周期刷新（R228A；本件无 TON） —— *)
rtReset(CLK := bReset);                                     // 复位沿 / Reset edge

(* —— 段 1：单拍/输出量预置（锁存量 _eCause/_bFault 不入清单，R107） —— *)
fOcvNormMv := 0.0;                                          // 归一值预置 / Normalised value preset
bInBand    := FALSE;                                        // 合格位预置 / In-band preset
eGrade     := E_DL_OtnGrade.eNoGrade;                       // 分级预置为"未分级" / Grade preset to ungraded
bValid     := FALSE;                                        // 有效性预置 / Validity preset
bClamped   := FALSE;                                        // 钳位标志预置 / Clamp flag preset
bError     := FALSE;                                        // 故障标志预清（R45 配对） / Error preset
_fNorm     := 0.0;                                          // 归一工作值预置 / Working value preset

(* —— 段 2：组态闸（合格带倒置 / 钳位限非正 → 故障锁存） —— *)
_bBandOk := (fBandLowMv < fBandHighMv);                     // 下限必须严格小于上限 / Lower must be strictly below upper
_fLim := fNormClampMv;                                      // 先直取脚值 / Take the pin value first
IF (NOT _bBandOk) OR (_fLim <= 0.0) OR (_fLim <> _fLim) OR ((_fLim - _fLim) <> (_fLim - _fLim)) THEN
    _fLim := DL_OTN_CLAMP_DEF;                              // 钳位限回退默认常量（与被判量解耦） / Fall back to the default limit
    _eCause := E_DL_OtnCause.eCfgIllegal;                   // 归因：组态非法 / Cause: illegal configuration
    _bFault := TRUE;                                        // 锁存 / Latch
    _eState := E_DL_OtnState.eFault;                        // 入故障相 / Enter fault phase
END_IF

(* —— 段 3：温度系数零闸（k=0 使归一恒等，判据静默失效，按故障处理 R179） —— *)
IF (_eState <> E_DL_OtnState.eFault) THEN
    IF (fTempCoeff = 0.0) OR (fTempCoeff <> fTempCoeff) OR ((fTempCoeff - fTempCoeff) <> (fTempCoeff - fTempCoeff)) THEN
        _eCause := E_DL_OtnCause.eCoeffZero;                // 归因：温度系数为零或非有限 / Cause: zero or non-finite coefficient
        _bFault := TRUE;                                    // 锁存 / Latch
        _eState := E_DL_OtnState.eFault;                    // 入故障相 / Enter fault phase
    END_IF
    IF (iTempUnit = E_DL_OtnUnit.eUnknown) THEN
        _eCause := E_DL_OtnCause.eUnitBad;                  // 归因：温度单位未知 / Cause: unknown temperature unit
        _bFault := TRUE;                                    // 锁存 / Latch
        _eState := E_DL_OtnState.eFault;                    // 入故障相 / Enter fault phase
    END_IF
END_IF

(* —— 段 4：迁出链（bReset 上升沿 → 待机相；解除式恒可达） —— *)
IF rtReset.Q THEN
    _bFault := FALSE;                                       // 清故障锁存 / Clear fault latch
    _eCause := E_DL_OtnCause.eNone;                         // 清成因 / Clear cause
    _eState := E_DL_OtnState.eIdle;                         // 回待机相 / Back to idle
END_IF

(* —— 段 5：相迁移（使能驱动；故障相由段 4 迁出） —— *)
CASE _eState OF

E_DL_OtnState.eIdle:
    IF bEnable THEN
        _eState := E_DL_OtnState.eRun;                      // 使能即进判据相 / Enable enters the running phase
    END_IF

E_DL_OtnState.eRun:
    IF NOT bEnable THEN
        _eState := E_DL_OtnState.eIdle;                     // 失能回待机相（不借故障相过桥，R211） / Disable returns to idle
    END_IF

E_DL_OtnState.eFault:
    ;                                                       // 故障相：由段 4 复位沿迁出 / Exit handled by the reset edge

ELSE
    _eCause := E_DL_OtnCause.ePhaseBad;                     // 归因：非法相位 / Cause: illegal phase
    _bFault := TRUE;                                        // 锁存 / Latch
    _eState := E_DL_OtnState.eFault;                        // 强拉故障相 / Force fault phase

END_CASE

(* —— 段 6：归一与判带（仅在判据相且样本有限时；非有限样本当拍不判、不锁存） —— *)
IF _eState = E_DL_OtnState.eRun THEN
    _bXFin := NOT ((fOcvMeasMv <> fOcvMeasMv) OR ((fOcvMeasMv - fOcvMeasMv) <> (fOcvMeasMv - fOcvMeasMv)))
          AND NOT ((fTempMeas <> fTempMeas) OR ((fTempMeas - fTempMeas) <> (fTempMeas - fTempMeas)))
          AND NOT ((fTempRefC <> fTempRefC) OR ((fTempRefC - fTempRefC) <> (fTempRefC - fTempRefC)));
    IF _bXFin THEN
        (* 单位换算（复用 FC_DL_TempUnitConvert 语义，三支全列、无 ELSE 猜默认） *)
        CASE iTempUnit OF
        E_DL_OtnUnit.eCelsius:
            _fTempC := fTempMeas;                           // 摄氏直通 / Celsius passes through
        E_DL_OtnUnit.eFahrenheit:
            _fTempC := (fTempMeas - DL_OTN_F_OFFS) * DL_OTN_F_SCALE;   // 华氏转摄氏 / Fahrenheit to Celsius
        E_DL_OtnUnit.eKelvin:
            _fTempC := fTempMeas - DL_OTN_K2C;               // 开尔文转摄氏 / Kelvin to Celsius
        ELSE
            _fTempC := fTempRefC;                           // 未知单位：取基准温度（段 3 已锁存故障，此支仅防未定义值）
        END_CASE

        _fNorm := fOcvMeasMv + fTempCoeff * (_fTempC - fTempRefC);      // 一阶线性归一 / First-order linear normalisation

        IF (_fNorm > _fLim) THEN
            _fNorm := _fLim;                                // 上钳 / Clamp high
            bClamped := TRUE;                               // 置钳位标志 / Raise the clamp flag
        ELSIF (_fNorm < (0.0 - _fLim)) THEN
            _fNorm := 0.0 - _fLim;                          // 下钳 / Clamp low
            bClamped := TRUE;                               // 置钳位标志 / Raise the clamp flag
        END_IF

        bValid := TRUE;                                     // 样本有限且已归一：结果有效 / Sample finite and normalised

        (* 判带（差值容差，禁 = 判等） *)
        IF ABS(_fNorm - fBandHighMv) < DL_OTN_EPS THEN
            eGrade := E_DL_OtnGrade.eHigh;                  // 贴上限：归高档（边界样本显式归属） / On the upper edge: graded high
            bInBand := TRUE;                                // 落在带内 / Inside the band
        ELSIF ABS(_fNorm - fBandLowMv) < DL_OTN_EPS THEN
            eGrade := E_DL_OtnGrade.eLow;                   // 贴下限：归低档 / On the lower edge: graded low
            bInBand := TRUE;                                // 落在带内 / Inside the band
        ELSIF _fNorm > fBandHighMv THEN
            eGrade := E_DL_OtnGrade.eHigh;                  // 超上限 / Above the upper limit
            bInBand := FALSE;                               // 带外 / Outside the band
        ELSIF _fNorm < fBandLowMv THEN
            eGrade := E_DL_OtnGrade.eLow;                   // 低于下限 / Below the lower limit
            bInBand := FALSE;                               // 带外 / Outside the band
        ELSE
            eGrade := E_DL_OtnGrade.eInBand;                // 严格带内 / Strictly inside the band
            bInBand := TRUE;                                // 合格 / Accept
        END_IF
    END_IF
END_IF

(* —— 段 7：出口单点映射（名实双出口，R191） —— *)
fOcvNormMv := _fNorm;                                       // 归一值出口（无效拍输出 0） / Normalised value outlet
eState     := _eState;                                      // 相出口 / Phase outlet
eCause     := _eCause;                                      // 成因出口 / Cause outlet
bError     := _bFault;                                      // 故障标志 / Error flag

END_FUNCTION_BLOCK

(* ---- FB_DL_PackHousingTighten.st ---- *)
(*==============================================================================
 * 组件名称 (Component)  : FB_DL_PackHousingTighten
 * 所属子库 (Sublibrary) : DL_Process
 * 当前版本 (Version)    : 1.0.0
 * 兼容性   (Platform)   : CODESYS 3.5+ / TwinCAT 3 / 汇川 InoProShop / 施耐德 Machine Expert
 *                         仅依赖 Standard.library（TON / R_TRIG），零厂商私有库
 * 功能描述 (Function)   : 电池包壳体螺栓拧紧对角轴序 + 扭矩/角度双窗判定。
 *                         ① 对角轴序：四螺栓按 1 → 3 → 2 → 4 的对角顺序拧（顺序常量表
 *                            DL_PTH_SEQ = [0, 2, 1, 3]），对角拧紧是为避免壳体单侧先压紧
 *                            导致密封面翘曲——顺序写死在常量里，不运行期可改。
 *                         ② 每一步由 bStepDone 上升沿推进（拧紧工具给"本颗完成"信号），
 *                            完成时即用该颗的 afTorque[i] / afAngle[i] 判双窗：
 *                            扭矩 ∈ [fTorqueLo, fTorqueHi] 且 角度 ∈ [fAngleLo, fAngleHi]，
 *                            任一越窗即该颗不合格。
 *                         ③ 不合格记录轴号：不合格螺栓的**螺栓号（1..4，非数组下标）**写入
 *                            anFailBolt 数组（按不合格先后排放），nFailCount 为个数。
 *                            记录轴号而不是只置一个 bNg，是因为返修要知道"回去拧哪一颗"。
 *                         ④ 四颗走完 → bCycleDone 单拍脉冲，bAllOk =（nFailCount = 0）。
 *                         ⑤ 每步有专用超时 tonStepTo（R228A 专用超时 TON 命名豁免），
 *                            超时 → eFault（eStepTimeout），记录卡住的螺栓号。
 * 接口     (Interface)  : 输入 afTorque / afAngle 四颗实测扭矩与角度（VAR_IN_OUT，本件只读）、
 *                         扭矩窗 fTorqueLo / fTorqueHi、角度窗 fAngleLo / fAngleHi、
 *                         bStart 启动沿、bStepDone 本颗完成沿、tStepTimeout 单颗超时、bReset 复位；
 *                         输出 nCurrentBolt 当前螺栓号（1..4，0=无）、bStepActive 拧紧进行中、
 *                         bCycleDone 一轮完成单拍、bAllOk 全合格、anFailBolt 不合格螺栓号表、
 *                         nFailCount 不合格个数、nDoneCount 已完成个数、eState / eCause / bError。
 * 边界     (Boundary)   : ① **属主边界（写死）：本件只排轴序与判双窗，不驱动拧紧轴、不下发扭矩
 *                         设定值、不做扭矩闭环**。工具动作与设定值下发属拧紧控制器/轴级 POU；
 *                         本件吃完成信号与实测值，出轴序推进与判定结论。
 *                         ② 组态闸：fTorqueLo <= 0.0、fTorqueHi <= fTorqueLo、fAngleLo < 0.0、
 *                         fAngleHi <= fAngleLo、tStepTimeout <= T#0S、任一实测 NaN
 *                         → 故障锁存（NaN 会让双窗比较恒假，静默判合格是最坏结果）。
 *                         ③ 固定四颗（ARRAY[0..3]）：颗数写死在类型里；若工艺要 6 颗须改类型与
 *                         顺序常量，不允许运行期可变（越界风险）。
 *                         ④ 单枚 TON（tonStepTo）+ 三枚 R_TRIG（bStart / bStepDone / bReset）
 *                         段 0 无条件周期刷新；tonStepTo 的 IN =（eRun 相），出相即复位，
 *                         不存在跨步累积（R228A）。
 *                         ⑤ eFault 迁出：bReset 上升沿 → eIdle（R228B）；另 bStart 上升沿亦可
 *                         从 eDone 重开一轮（新工件，非解除式）。
 *                         ⑥ 零全局耦合（无 GVL / 无 VAR_EXTERNAL / 无物理地址）。
 * 分工声明 (Scope)      : 与 `FB_DL_AxisTorqueLimitGuard`（轴力矩瞬时限）分工——那件是运动中
 *                         连续保护，本件是**工序级**顺序与结果判定；不共用判据、不互相内嵌。
 * 来源标签 (Source Tag) : ROADMAP B 类 / T2-2（电池包壳体螺栓对角拧紧，自研 clean-room）
 * 解除式   (Release)    : bReset 上升沿 ∧ 组态合法 → 清故障、清不合格表、回 eIdle。
 *                         自证可满足：复位为外部动作，无锁存量门控。
 * 码表     (Codes)      : 本件不占用任何全局数字码位。出口为 INT 螺栓号 + INT 表 + BOOL 组 +
 *                         ENUM（eState / eCause）；数字码位待主控收口阶段统一派号。
 * 红线自检 (Redline)    : R1 ✓ 零 GVL/VAR_EXTERNAL ｜ R2 ✓ 零 %I/%Q/%M ｜ R3 ✓ 纯 IEC 61131-3
 *                         R4 ✓ 数组边界闸 + 双窗几何闸 + NaN 闸 ｜ R5 ✓ 声明逐行同行双语注释
 *                         R6 ✓ ENUM+CASE 含 ELSE ｜ R7 ✓ TON/R_TRIG 段 0 无条件刷新
 * 修订历史 (Revision)   : 2026-11-19  v1.0.0  R46 首版（批次 4 · 序号 20）
 *==============================================================================*)

TYPE E_DL_PthState :
(
    eIdle  := 0,    // 待启动 / Idle
    eRun   := 10,   // 拧紧进行相（逐颗推进） / Tightening, advancing bolt by bolt
    eDone  := 20,   // 一轮完成相（结论已出） / Cycle complete with a verdict
    eFault := 90    // 故障相（超时/组态非法，等复位） / Fault, awaiting reset
);
END_TYPE

TYPE E_DL_PthCause :
(
    eNone        := 0,   // 无异常 / No anomaly
    eCfgIllegal  := 1,   // 组态非法（窗口倒置/超时非正/实测非有限） / Illegal configuration
    eTorqueNg    := 2,   // 扭矩越窗 / Torque out of the window
    eAngleNg     := 3,   // 角度越窗 / Angle out of the window
    eBothNg      := 4,   // 扭矩与角度同时越窗 / Torque and angle both out of the window
    eStepTimeout := 5,   // 单颗拧紧超时 / Single-bolt tightening timed out
    ePhaseBad    := 6    // 非法相位兜底 / Illegal phase fallback
);
END_TYPE

FUNCTION_BLOCK FB_DL_PackHousingTighten
VAR_IN_OUT
    afTorque : ARRAY[0..3] OF REAL;     // 四颗实测扭矩（本件只读） [N·m] / Four measured torques, read-only here [N·m]
    afAngle  : ARRAY[0..3] OF REAL;     // 四颗实测转角（本件只读） [度] / Four measured angles, read-only here [deg]
END_VAR
VAR_INPUT
    fTorqueLo    : REAL := 20.0;        // 扭矩窗下限，域 > 0.0 [N·m] / Torque window lower limit, > 0.0 [N·m]
    fTorqueHi    : REAL := 30.0;        // 扭矩窗上限，域 > fTorqueLo [N·m] / Torque window upper limit, > lower [N·m]
    fAngleLo     : REAL := 10.0;        // 角度窗下限，域 >= 0.0 [度] / Angle window lower limit, >= 0.0 [deg]
    fAngleHi     : REAL := 90.0;        // 角度窗上限，域 > fAngleLo [度] / Angle window upper limit, > lower [deg]
    bStart       : BOOL := FALSE;       // 启动沿，开新的一轮 [-] / Start edge, opens a new cycle
    bStepDone    : BOOL := FALSE;       // 本颗拧紧完成沿，推进一颗 [-] / Current-bolt-done edge, advances one bolt
    tStepTimeout : TIME := T#10S;       // 单颗超时，域 > T#0S [ms] / Per-bolt timeout, > T#0S [ms]
    bReset       : BOOL := FALSE;       // 复位，上升沿清故障与不合格表 [-] / Reset, clears fault and the failure table
END_VAR
VAR_OUTPUT
    nCurrentBolt : INT;                 // 当前螺栓号 1..4，0=无 [号] / Current bolt number, 1..4, 0 means none
    bStepActive  : BOOL;                // 拧紧进行中（有当前螺栓） [-] / Tightening in progress
    bCycleDone   : BOOL;                // 一轮完成，单拍脉冲 [-] / Cycle done, single-scan pulse
    bAllOk       : BOOL;                // 本轮全合格 [-] / All bolts passed this cycle
    anFailBolt   : ARRAY[0..3] OF INT;  // 不合格螺栓号表（按发生先后，0 表空位） [号] / Failed bolt numbers in order, 0 marks an empty slot
    nFailCount   : INT;                 // 不合格个数 [颗] / Number of failed bolts
    nDoneCount   : INT;                 // 已完成颗数 [颗] / Number of completed bolts
    eState       : E_DL_PthState;       // 状态出口 [-] / State outlet
    eCause       : E_DL_PthCause;       // 成因出口（R190 归因唯一） [-] / Cause outlet
    bError       : BOOL;                // 故障标志（超时/组态非法） [-] / Error flag
END_VAR
VAR
    _eState    : E_DL_PthState := E_DL_PthState.eIdle;    // 内部相位（CASE 唯一写入目标） / Internal phase
    _eCause    : E_DL_PthCause := E_DL_PthCause.eNone;    // 成因锁存量 / Latched cause
    tonStepTo  : TON;           // 单颗拧紧专用超时，段 0 无条件调用 / Per-bolt dedicated timeout
    rtStart    : R_TRIG;        // 启动沿实例，段 0 无条件调用 / Start edge instance
    rtStepDone : R_TRIG;        // 本颗完成沿实例，段 0 无条件调用 / Step-done edge instance
    rtReset    : R_TRIG;        // 复位沿实例，段 0 无条件调用 / Reset edge instance
    _nStepIdx  : INT;           // 顺序表下标 0..3（锁存量） / Sequence table index, latched
    _nFailCnt  : INT;           // 不合格计数（锁存量） [颗] / Failure count, latched
    _nDoneCnt  : INT;           // 完成计数（锁存量） [颗] / Done count, latched
    _anFail    : ARRAY[0..3] OF INT;    // 不合格螺栓号表（锁存量） [号] / Failure table, latched
    _bFault    : BOOL;          // 故障锁存位（锁存量） / Latched fault bit
    _bCfgBad   : BOOL;          // 组态非法当拍量 [-] / Illegal configuration this scan
    _bNonFin   : BOOL;          // 实测非有限当拍量 [-] / Non-finite measurement this scan
    _bTqNg     : BOOL;          // 当前颗扭矩越窗当拍量 [-] / Torque NG for the current bolt
    _bAgNg     : BOOL;          // 当前颗角度越窗当拍量 [-] / Angle NG for the current bolt
    _nIdxSafe  : INT;           // 钳位后的顺序表下标（0..3） / Clamped sequence index
    _i         : INT;           // 遍历索引 / Loop index
END_VAR
VAR CONSTANT
    DL_PTH_N       : INT := 4;                          // 螺栓颗数（与 ARRAY 上界一致） [颗] / Bolt count matching the array bounds
    DL_PTH_SEQ     : ARRAY[0..3] OF INT := [0, 2, 1, 3];    // 对角顺序表：1→3→2→4（0 基下标） [下标] / Diagonal order 1-3-2-4 as 0-based indices
END_VAR

(* —— 段 0：组态闸派生 + 四实例无条件周期刷新 —— *)
_bNonFin := FALSE;                                                  // 非有限标志初值 / Non-finite initial value
FOR _i := 0 TO DL_PTH_N - 1 DO
    IF (afTorque[_i] <> afTorque[_i]) OR (afAngle[_i] <> afAngle[_i]) THEN
        _bNonFin := TRUE;                                           // 实测 NaN 自反判（判等禁令唯一例外） / Measurement NaN test
    END_IF
END_FOR
_bCfgBad := (fTorqueLo <= 0.0) OR (fTorqueHi <= fTorqueLo)          // 扭矩窗几何闸 / Torque window geometry
         OR (fAngleLo < 0.0) OR (fAngleHi <= fAngleLo)              // 角度窗几何闸 / Angle window geometry
         OR (tStepTimeout <= T#0S) OR _bNonFin;                     // 超时闸 + 非有限 / Timeout gate and non-finite
rtStart(CLK := bStart);                                             // 启动沿，每拍必调（R228A） / Start edge, every scan
rtStepDone(CLK := bStepDone);                                       // 完成沿，每拍必调 / Step-done edge, every scan
rtReset(CLK := bReset);                                             // 复位沿，每拍必调 / Reset edge, every scan
tonStepTo(IN := (_eState = E_DL_PthState.eRun), PT := tStepTimeout);    // 单颗专用超时（进相计时，出相自复位） / Per-bolt dedicated timeout

(* —— 段 1：单拍量预清零（锁存量 _nStepIdx/_nFailCnt/_nDoneCnt/_anFail/_bFault 不入清单，R107） —— *)
bCycleDone  := FALSE;           // 完成脉冲预清 / Cycle-done preset
bStepActive := FALSE;           // 进行中指示预清 / Step-active preset
bAllOk      := FALSE;           // 全合格位预清 / All-ok preset
bError      := FALSE;           // 故障标志预清（R45 配对） / Error flag preset
_bTqNg      := FALSE;           // 扭矩越窗当拍量预清 / Torque NG preset
_bAgNg      := FALSE;           // 角度越窗当拍量预清 / Angle NG preset

(* —— 段 2：复位沿（清故障、清表、回待机） —— *)
IF rtReset.Q THEN
    _bFault   := FALSE;                                 // 清故障锁存 / Clear the fault latch
    _eCause   := E_DL_PthCause.eNone;                   // 清成因 / Clear cause
    _nFailCnt := 0;                                     // 不合格计数清零 / Failure count cleared
    _nDoneCnt := 0;                                     // 完成计数清零 / Done count cleared
    _nStepIdx := 0;                                     // 顺序下标归零 / Sequence index cleared
    FOR _i := 0 TO DL_PTH_N - 1 DO
        _anFail[_i] := 0;                               // 不合格表清零 / Failure table cleared
    END_FOR
    IF _eState <> E_DL_PthState.eIdle THEN
        _eState := E_DL_PthState.eIdle;                 // 回待机相（R228B 迁出路径） / Back to idle, the R228B exit
    END_IF
END_IF
IF _bCfgBad THEN
    _bFault := TRUE;                                    // 组态非法锁存 / Latch illegal configuration
    _eCause := E_DL_PthCause.eCfgIllegal;               // 归因：组态非法 / Cause: illegal configuration
    _eState := E_DL_PthState.eFault;                    // 入故障相 / Enter fault phase
END_IF

(* —— 段 3：启动沿（开新的一轮，清表清计数） —— *)
IF rtStart.Q AND (NOT _bCfgBad) THEN
    _nStepIdx := 0;                                     // 从顺序表第 0 位开始 / Start at sequence position 0
    _nFailCnt := 0;                                     // 不合格计数清零 / Failure count cleared
    _nDoneCnt := 0;                                     // 完成计数清零 / Done count cleared
    FOR _i := 0 TO DL_PTH_N - 1 DO
        _anFail[_i] := 0;                               // 表清零（新工件） / Table cleared for the new part
    END_FOR
    _eCause   := E_DL_PthCause.eNone;                   // 清成因 / Clear cause
    _eState   := E_DL_PthState.eRun;                    // 入运行相 / Enter run phase
END_IF

(* —— 段 4：逐颗推进与双窗判定（完成沿触发，单点写入锁存量，R187） —— *)
IF (_eState = E_DL_PthState.eRun) AND rtStepDone.Q AND (NOT _bCfgBad) THEN
    _nIdxSafe := _nStepIdx;                             // 取顺序下标 / Take the sequence index
    IF _nIdxSafe < 0 THEN
        _nIdxSafe := 0;                                 // 下界钳（双保险） / Lower clamp
    END_IF
    IF _nIdxSafe > DL_PTH_N - 1 THEN
        _nIdxSafe := DL_PTH_N - 1;                      // 上界钳（双保险，绝不越 ARRAY） / Upper clamp, never index past the array
    END_IF
    _bTqNg := (afTorque[DL_PTH_SEQ[_nIdxSafe]] < fTorqueLo) OR (afTorque[DL_PTH_SEQ[_nIdxSafe]] > fTorqueHi);    // 扭矩双窗 / Torque window, both sides
    _bAgNg := (afAngle[DL_PTH_SEQ[_nIdxSafe]] < fAngleLo) OR (afAngle[DL_PTH_SEQ[_nIdxSafe]] > fAngleHi);       // 角度双窗 / Angle window, both sides
    IF _bTqNg OR _bAgNg THEN
        IF _nFailCnt < DL_PTH_N THEN
            _anFail[_nFailCnt] := DL_PTH_SEQ[_nIdxSafe] + 1;    // 记录螺栓号（1 基，不是数组下标） / Record the 1-based bolt number
            _nFailCnt := _nFailCnt + 1;                         // 计数增 / Increment the count
        END_IF
        IF _bTqNg AND _bAgNg THEN
            _eCause := E_DL_PthCause.eBothNg;                   // 归因：双窗同越 / Cause: both windows violated
        ELSIF _bTqNg THEN
            _eCause := E_DL_PthCause.eTorqueNg;                 // 归因：扭矩越窗 / Cause: torque violated
        ELSE
            _eCause := E_DL_PthCause.eAngleNg;                  // 归因：角度越窗 / Cause: angle violated
        END_IF
    END_IF
    _nDoneCnt := _nDoneCnt + 1;                                 // 完成颗数增 / Increment the done count
    _nStepIdx := _nStepIdx + 1;                                 // 顺序推进 / Advance the sequence
    IF _nStepIdx >= DL_PTH_N THEN
        _eState := E_DL_PthState.eDone;                         // 四颗走完：出结论 / All four done, deliver the verdict
        bCycleDone := TRUE;                                     // 单拍完成脉冲 / Single-scan completion pulse
    END_IF
END_IF

(* —— 段 5：单颗超时（运行相且计时到 → 故障，记录卡住的螺栓号） —— *)
IF (_eState = E_DL_PthState.eRun) AND tonStepTo.Q AND (NOT _bCfgBad) THEN
    IF _nFailCnt < DL_PTH_N THEN
        _nIdxSafe := _nStepIdx;                                 // 取当前下标 / Take the present index
        IF _nIdxSafe < 0 THEN
            _nIdxSafe := 0;                                     // 下界钳 / Lower clamp
        END_IF
        IF _nIdxSafe > DL_PTH_N - 1 THEN
            _nIdxSafe := DL_PTH_N - 1;                          // 上界钳 / Upper clamp
        END_IF
        _anFail[_nFailCnt] := DL_PTH_SEQ[_nIdxSafe] + 1;        // 记录超时螺栓号 / Record the timed-out bolt number
        _nFailCnt := _nFailCnt + 1;                             // 计数增 / Increment the count
    END_IF
    _bFault := TRUE;                                            // 锁存 / Latch
    _eCause := E_DL_PthCause.eStepTimeout;                      // 归因：单颗超时 / Cause: per-bolt timeout
    _eState := E_DL_PthState.eFault;                            // 入故障相 / Enter fault phase
END_IF

(* —— 段 6：锁存相位迁移闸 —— *)
IF _bFault AND (_eState <> E_DL_PthState.eFault) THEN
    _eState := E_DL_PthState.eFault;                            // 锁存即入故障相 / Latch enters fault phase
END_IF

(* —— 段 7：相位机（ENUM 全成员显式标签 + ELSE 兜底，R128） —— *)
CASE _eState OF

E_DL_PthState.eIdle:
    IF _bCfgBad THEN                                            // 出口 1：组态非法 / Illegal configuration
        _eState := E_DL_PthState.eFault;
    ELSIF rtStart.Q THEN                                        // 出口 2：启动沿 / Start edge
        _eState := E_DL_PthState.eRun;
    END_IF

E_DL_PthState.eRun:
    IF _bCfgBad OR _bFault THEN                                 // 出口 1：故障（组态或超时） / Fault, config or timeout
        _eState := E_DL_PthState.eFault;
    ELSIF _nStepIdx >= DL_PTH_N THEN                            // 出口 2：四颗走完 / All four finished
        _eState := E_DL_PthState.eDone;
    END_IF

E_DL_PthState.eDone:
    IF _bCfgBad THEN                                            // 出口 1：组态非法 / Illegal configuration
        _eState := E_DL_PthState.eFault;
    ELSIF rtStart.Q THEN                                        // 出口 2：新工件启动 / New part started
        _eState := E_DL_PthState.eRun;
    END_IF

E_DL_PthState.eFault:
    IF rtReset.Q AND (NOT _bCfgBad) THEN                        // 出口：复位且组态已合法才迁出（R228B） / Reset with legal config
        _eState := E_DL_PthState.eIdle;
    END_IF

ELSE
    _eCause := E_DL_PthCause.ePhaseBad;                         // 归因：非法相位 / Cause: illegal phase
    _eState := E_DL_PthState.eFault;                            // 强拉故障相 / Force fault phase
    bError  := TRUE;                                            // 故障标志 / Error flag

END_CASE

(* —— 段 8：出口单点映射（当前螺栓号由顺序表反查，1 基；名实双出口 R191） —— *)
nCurrentBolt := 0;                                              // 当前螺栓号缺省无 / Current bolt defaults to none
IF _eState = E_DL_PthState.eRun THEN
    _nIdxSafe := _nStepIdx;                                     // 取顺序下标 / Take the sequence index
    IF _nIdxSafe < 0 THEN
        _nIdxSafe := 0;                                         // 下界钳 / Lower clamp
    END_IF
    IF _nIdxSafe > DL_PTH_N - 1 THEN
        _nIdxSafe := DL_PTH_N - 1;                              // 上界钳 / Upper clamp
    END_IF
    nCurrentBolt := DL_PTH_SEQ[_nIdxSafe] + 1;                  // 螺栓号 1..4（对角序反查） / Bolt number 1..4 via the diagonal order
END_IF
bStepActive := (_eState = E_DL_PthState.eRun) AND (nCurrentBolt > 0);      // 进行中 = 运行相且有当前螺栓 / Active when running with a current bolt
bAllOk      := (_eState = E_DL_PthState.eDone) AND (_nFailCnt = 0);        // 全合格 = 完成相且无不合格 / All-ok when done with no failures
nFailCount  := _nFailCnt;                                       // 不合格个数出口 / Failure count outlet
nDoneCount  := _nDoneCnt;                                       // 完成颗数出口 / Done count outlet
FOR _i := 0 TO DL_PTH_N - 1 DO
    anFailBolt[_i] := _anFail[_i];                              // 不合格表整体回放 / Failure table replay
END_FOR
bError := _bFault OR _bCfgBad;                                  // 故障标志 = 锁存或组态非法 / Error = latch or illegal config
eState := _eState;                                              // 状态出口 / State outlet
eCause := _eCause;                                              // 成因出口 / Cause outlet

END_FUNCTION_BLOCK

(* ---- FB_DL_PackMlStateMachine.st ---- *)
(*==============================================================================
 * 组件名称 (Component)  : FB_DL_PackMlStateMachine
 * 所属子库 (Sublibrary) : DL_Process
 * 当前版本 (Version)    : 1.0.0
 * 组件分类 (Category)   : 功能块（FUNCTION_BLOCK）· PackML 状态机框架 · Level 2 机台层
 * 兼容性   (Platform)   : CODESYS 3.5 / TwinCAT 3 / 汇川 InoProShop / Schneider
 *                         Machine Expert；仅依赖 Standard.library，零厂商方言
 * 功能描述 (Function)   : PackML / ISA-TR88.00.02 十七态（+ Undefined 占位）
 *                         状态机 clean-room 框架实现。命令驱动 + acting 态由
 *                         bStateComplete 自动推进；本块不编排任何具体工艺
 *                         动作——纯状态机框架，动作由调用方按态派发（Level 2
 *                         依赖注入原则），与机台工艺完全解耦。
 * 设计要点 (Key notes)  : ① Aborting 为最高优先级出口：bProcessAbort 或非法态
 *                           → eAborting（CASE+ELSE 兜底同向，公约 0.1/0.2）；
 *                         ② Clearing 完成后必经 eStopped（S-1「abort 后强制
 *                           去污步」语义）；Aborted 恢复链 Clear→Clearing→
 *                           Stopped→Reset→Resetting→Idle；
 *                         ③ eExecute 中 bInterlockOk 失失 → 自动转 eHolding
 *                           （机内保持），与 eSuspended（机外挂起）区分指示，
 *                           保 OEE 根因数据质量（S-1 提取点⑤）；
 *                         ④ 模式切换仅允许 eStopped/eIdle/eCompleted 稳态
 *                           （S-1 提取点⑥），其余态下变更被拒并置信息级
 *                           0005_0101；
 *                         ⑤ 首扫/跟踪判据唯一合法范式 IF bTrack OR (NOT bInit)
 *                           （公约 0.1）：首扫从 eUndefined 迁入 eStopped，
 *                           运行中途跟踪脉冲不扰动已建立的状态；
 *                         ⑥ ePrevState 仅在真实跃迁时刷新，Abort 路径保留
 *                           跃迁前状态供 HMI 复盘。
 * 枚举归属 (Enum note)  : E_DL_PackMlState / E_DL_PackMlCmd / E_DL_UnitMode
 *                         三个 DUT 随本块同文件发布（规格书第 6 节交付约定），
 *                         FB_DL_PackMlCmdDecoder 引用 E_DL_PackMlCmd，导入
 *                         本文件后全局可见。
 * 开源溯源 (Origin)     : packml。来源为 OMAC PackML / ISA-TR88.00.02 公开
 *                         规范的状态集合、命令集合与跃迁语义（S-1 提取点
 *                         ①②③④⑤⑥），状态编号逐项对齐；实现与命名 100%
 *                         自有 clean-room，不参考任何厂商 LUC 代码结构。
 * 验收向量 (Acceptance) :
 *   V1 正常链：eIdle → Start → eStarting →(SC)→ eExecute → Complete →
 *      eCompleting →(SC)→ eCompleted → Reset → eResetting →(SC)→ eIdle；
 *   V2 Abort→Clear→Reset 全恢复链：任意态 bProcessAbort → eAborting →
 *      eAborted → Clear → eClearing →(SC)→ eStopped → Reset → eIdle；
 *   V3 非法态兜底：强制 _eState=88 → ELSE 兜底 → eAborting，码 0005_0201；
 *   V4 非稳态模式切换：eExecute 下改 eMode → 拒绝 + 信息级 0005_0101；
 *   V5 联锁失失保持：eExecute 中 bInterlockOk=FALSE → eHolding，
 *      bHeldByMachine=TRUE；Unhold → eUnholding →(SC)→ eExecute；
 *   V6 中途跟踪脉冲：eExecute 中 bTrack=TRUE 一拍 → 状态保持不扰动。
 * 故障码表 (Error codes):
 *   16#0005_0101【信息级】非稳态模式切换被拒 / 16#0005_0201【故障级】
 *   非法状态兜底（走 Aborting 路径）。
 * 修订历史 (Revision)   :
 *   2026-11-15  v1.0.0  首版入库（Round 05 · DL_Process 立项）
 *============================================================================*)

(*-----------------------------------------------------------------------------
 * 调用示例 (Instance guide)：
 *   fbPml.eMode := E_DL_PackMlMode.eProduction;   // 组态期或稳态期切换
 *   fbPml.eCmd := fbDecoder.eCmd;                 // 命令由解码器单发供给
 *   fbPml(bStateComplete := fbStep.bSeqDone,      // 周期调用
 *         bInterlockOk := bSafeChain, bProcessAbort := bEstopChain);
 *   工艺派发示例：按 fbPml.eState 分态派发，eExecute 态执行 fbStation.Run()。
 *   OEE 采集：bInExecute 计 Execute 时长；bHeldByMachine/bSuspendedByLine
 *   分别归因机内保持与机外挂起，根因统计勿混用。
 *----------------------------------------------------------------------------*)

{attribute 'strict'}
{attribute 'qualified_only'}
TYPE E_DL_PackMlState :
(
    eUndefined    := 0,    // 未定义：上电占位态，首扫迁移至 eStopped / Undefined: power-up placeholder, migrated at first scan
    eClearing     := 1,    // 清除中（acting，自动推进）：abort 后强制去污步 / Clearing (acting): mandatory cleanup after abort
    eStopped      := 2,    // 已停止（wait）：复位/启动/急停出口 / Stopped (wait): reset, start or abort exits
    eStarting     := 3,    // 启动中（acting，自动推进）：预热/自检等启动子工序 / Starting (acting): startup sub-operations
    eIdle         := 4,    // 空闲（wait）：就绪待命，Start 进入生产 / Idle (wait): ready, Start enters production
    eSuspended    := 5,    // 已挂起（wait）：机外原因暂停（线体/供料） / Suspended (wait): paused by external line reason
    eExecute      := 6,    // 执行中（wait，生产主态）：工艺动作派发与 OEE 计时态 / Execute (wait): main production state for OEE
    eStopping     := 7,    // 停止中（acting，自动推进）：受控停机子工序 / Stopping (acting): controlled stop sub-operations
    eAborting     := 8,    // 急停中（acting，自动跃迁）：最高优先级出口 / Aborting (acting): highest-priority exit
    eAborted      := 9,    // 已急停（wait）：仅 Clear/Reset 可退 / Aborted (wait): only Clear or Reset exits
    eHolding      := 10,   // 保持中（acting，自动推进）：机内原因保持过渡态 / Holding (acting): machine-internal hold transition
    eHeld         := 11,   // 已保持（wait）：机内原因暂停，Unhold 恢复 / Held (wait): held by machine reason, Unhold resumes
    eUnholding    := 12,   // 恢复中（acting，自动推进）：从保持回到执行 / Unholding (acting): resuming from held
    eSuspending   := 13,   // 挂起中（acting，自动推进）：机外暂停过渡 / Suspending (acting): external suspend transition
    eUnsuspending := 14,   // 解挂中（acting，自动推进）：从挂起回到执行 / Unsuspending (acting): resuming from suspended
    eResetting    := 15,   // 复位中（acting，自动推进）：回 Idle 的复位子工序 / Resetting (acting): reset sub-operations to idle
    eCompleting   := 16,   // 完成中（acting，自动推进）：完工收尾子工序 / Completing (acting): completion sub-operations
    eCompleted    := 17    // 已完成（wait）：批次完成，Reset/Clear 退出 / Completed (wait): batch done, Reset or Clear exits
) UINT;
END_TYPE

{attribute 'strict'}
{attribute 'qualified_only'}
TYPE E_DL_PackMlCmd :
(
    eUndefined     := 0,   // 无命令占位（No command placeholder）
    eReset         := 1,   // 复位命令（Reset command）
    eStart         := 2,   // 启动命令（Start command）
    eStop          := 3,   // 停止命令（Stop command）
    eHold          := 4,   // 保持命令（Hold command）
    eUnhold        := 5,   // 解除保持命令（Unhold command）
    eSuspend       := 6,   // 挂起命令（Suspend command）
    eUnsuspend     := 7,   // 解除挂起命令（Unsuspend command）
    eAbort         := 8,   // 急停命令（Abort command）
    eClear         := 9,   // 清除命令（Clear command）
    eComplete      := 10,  // 完工命令（Complete command）
    eStateComplete := 11   // 子工序完成命令（State complete command），命令形态的 SC
) UINT;
END_TYPE

{attribute 'strict'}
{attribute 'qualified_only'}
TYPE E_DL_UnitMode :
(
    eInvalid     := 0,    // 无效模式占位（Invalid mode placeholder）
    eProduction  := 1,    // 生产模式（Production mode）
    eMaintenance := 2,    // 维护模式（Maintenance mode）
    eManual      := 3,    // 手动模式（Manual mode）
    eUser4       := 4,    // 用户自定义模式 4（User defined mode 4）
    eUser5       := 5,    // 用户自定义模式 5（User defined mode 5）
    eUser6       := 6,    // 用户自定义模式 6（User defined mode 6）
    eUser7       := 7,    // 用户自定义模式 7（User defined mode 7）
    eUser8       := 8,    // 用户自定义模式 8（User defined mode 8）
    eUser9       := 9,    // 用户自定义模式 9（User defined mode 9）
    eUser10      := 10,   // 用户自定义模式 10（User defined mode 10）
    eUser11      := 11,   // 用户自定义模式 11（User defined mode 11）
    eUser12      := 12,   // 用户自定义模式 12（User defined mode 12）
    eUser13      := 13,   // 用户自定义模式 13（User defined mode 13）
    eUser14      := 14,   // 用户自定义模式 14（User defined mode 14）
    eUser15      := 15    // 用户自定义模式 15（User defined mode 15）
) UINT;
END_TYPE

FUNCTION_BLOCK FB_DL_PackMlStateMachine
VAR_INPUT
    eMode          : E_DL_UnitMode := E_DL_UnitMode.eInvalid;      // 单元模式（Unit mode），S-1 提取点④，仅稳态可切换
    eCmd           : E_DL_PackMlCmd := E_DL_PackMlCmd.eUndefined;  // 标准命令（Standard command），由 FB_DL_PackMlCmdDecoder 单发供给
    bStateComplete : BOOL := FALSE;       // 子工序完成信号（State complete），acting 态推进用
    bInterlockOk   : BOOL := TRUE;        // 工艺联锁（Process interlock），Execute 态保持条件，失失转机内保持
    bProcessAbort  : BOOL := FALSE;       // 工艺级急停触发（Process abort trigger），如安全门/急停链，电平生效
    bTrack         : BOOL := FALSE;       // 跟踪脉冲（Tracking pulse），首扫/跟踪同步（R5 公约 0.1）
END_VAR
VAR_OUTPUT
    eState         : E_DL_PackMlState := E_DL_PackMlState.eUndefined;   // 当前状态（Current state）
    ePrevState     : E_DL_PackMlState := E_DL_PackMlState.eUndefined;   // 前一状态（Previous state），Abort 路径复盘用
    bInExecute     : BOOL := FALSE;       // Execute 态指示（In execute），OEE 计时用
    bHeldByMachine : BOOL := FALSE;       // 机内保持指示（Held by machine），OEE 根因：机内原因
    bSuspendedByLine : BOOL := FALSE;     // 机外挂起指示（Suspended by line），OEE 根因：机外原因
    uErrorId       : UDINT := 0;          // 末次事件码（Last error code），信息级码不构成故障
END_VAR
VAR
    bInit          : BOOL := FALSE;       // 首扫标志（First-scan flag，R19 范式配套）
    _eState        : E_DL_PackMlState := E_DL_PackMlState.eUndefined;   // 内部当前状态（Internal current state）
    _eStateOld     : E_DL_PackMlState := E_DL_PackMlState.eUndefined;   // 本拍跃迁前快照（Pre-transition snapshot）
    _ePrevState    : E_DL_PackMlState := E_DL_PackMlState.eUndefined;   // 内部前一状态（Internal previous state）
    _eModeActive   : E_DL_UnitMode := E_DL_UnitMode.eInvalid;           // 生效单元模式（Active unit mode），非稳态拒绝切换
    _eModeReqLast  : E_DL_UnitMode := E_DL_UnitMode.eInvalid;           // 上一拍模式请求（Last mode request），模式变更沿检测
END_VAR

// 段 1｜R19 首扫/跟踪同步：判据唯一合法范式 IF bTrack OR (NOT bInit)
IF bTrack OR (NOT bInit) THEN
    IF _eState = E_DL_PackMlState.eUndefined THEN
        _eState := E_DL_PackMlState.eStopped;          // PackML 上电默认稳态：Stopped
        _ePrevState := E_DL_PackMlState.eUndefined;
        _eModeActive := eMode;                         // 首扫锁定当前模式请求
    END_IF
    bInit := TRUE;                                     // 运行中途跟踪脉冲不扰动已建立状态（验收向量 V6）
END_IF

// 段 2｜工艺级急停最高优先级出口：任何非 Aborting/Aborted 态直达 eAborting
IF bProcessAbort AND (_eState <> E_DL_PackMlState.eAborting) AND (_eState <> E_DL_PackMlState.eAborted) THEN
    _ePrevState := _eState;                            // 保留跃迁前状态供 HMI 复盘
    _eState := E_DL_PackMlState.eAborting;
END_IF

// 段 3｜模式切换稳态门禁（S-1 提取点⑥）：仅 eStopped/eIdle/eCompleted 允许
IF eMode <> _eModeReqLast THEN                      // 新模式请求沿
    _eModeReqLast := eMode;
    IF (_eState = E_DL_PackMlState.eStopped) OR (_eState = E_DL_PackMlState.eIdle)
       OR (_eState = E_DL_PackMlState.eCompleted) THEN
        _eModeActive := eMode;                      // 稳态允许切换
    ELSE
        uErrorId := 16#0005_0101;                   // 信息级：非稳态模式切换被拒（R21：不置故障）
    END_IF
END_IF

// 段 4｜十七态主状态机：命令驱动 + acting 态 bStateComplete 自动推进
_eStateOld := _eState;                              // 跃迁前快照，供 ePrevState 刷新
CASE _eState OF

    E_DL_PackMlState.eUndefined:                    // 防御驻留态：首扫已迁移，非法驻留即回 Stopped
        _eState := E_DL_PackMlState.eStopped;

    E_DL_PackMlState.eClearing:                     // acting：清除进行中（abort 后强制去污步）
        IF bStateComplete OR (eCmd = E_DL_PackMlCmd.eStateComplete) THEN
            _eState := E_DL_PackMlState.eStopped;   // S-1：清除完成必经 Stopped
        END_IF

    E_DL_PackMlState.eStopped:                      // wait：复位/启动/急停出口
        IF eCmd = E_DL_PackMlCmd.eReset THEN
            _eState := E_DL_PackMlState.eResetting;
        ELSIF eCmd = E_DL_PackMlCmd.eStart THEN
            _eState := E_DL_PackMlState.eStarting;
        ELSIF eCmd = E_DL_PackMlCmd.eAbort THEN
            _eState := E_DL_PackMlState.eAborting;
        END_IF

    E_DL_PackMlState.eStarting:                     // acting：启动子工序（预热/自检等）
        IF bStateComplete OR (eCmd = E_DL_PackMlCmd.eStateComplete) THEN
            _eState := E_DL_PackMlState.eIdle;      // 启动完成回空闲
        END_IF

    E_DL_PackMlState.eIdle:                         // wait：就绪待命
        IF eCmd = E_DL_PackMlCmd.eStart THEN
            _eState := E_DL_PackMlState.eStarting;
        ELSIF eCmd = E_DL_PackMlCmd.eStop THEN
            _eState := E_DL_PackMlState.eStopping;
        ELSIF eCmd = E_DL_PackMlCmd.eAbort THEN
            _eState := E_DL_PackMlState.eAborting;
        END_IF

    E_DL_PackMlState.eSuspended:                    // wait：机外原因暂停
        IF eCmd = E_DL_PackMlCmd.eUnsuspend THEN
            _eState := E_DL_PackMlState.eUnsuspending;
        ELSIF eCmd = E_DL_PackMlCmd.eStop THEN
            _eState := E_DL_PackMlState.eStopping;
        ELSIF eCmd = E_DL_PackMlCmd.eAbort THEN
            _eState := E_DL_PackMlState.eAborting;
        END_IF

    E_DL_PackMlState.eExecute:                      // wait：生产主态，工艺动作由此派发
        IF NOT bInterlockOk THEN
            _eState := E_DL_PackMlState.eHolding;   // 联锁失失 → 机内保持（OEE 根因：机内）
        ELSIF bStateComplete OR (eCmd = E_DL_PackMlCmd.eStateComplete) OR (eCmd = E_DL_PackMlCmd.eComplete) THEN
            _eState := E_DL_PackMlState.eCompleting;
        ELSIF eCmd = E_DL_PackMlCmd.eHold THEN
            _eState := E_DL_PackMlState.eHolding;
        ELSIF eCmd = E_DL_PackMlCmd.eSuspend THEN
            _eState := E_DL_PackMlState.eSuspending;
        ELSIF eCmd = E_DL_PackMlCmd.eStop THEN
            _eState := E_DL_PackMlState.eStopping;
        ELSIF eCmd = E_DL_PackMlCmd.eAbort THEN
            _eState := E_DL_PackMlState.eAborting;
        END_IF

    E_DL_PackMlState.eStopping:                     // acting：受控停机子工序
        IF bStateComplete OR (eCmd = E_DL_PackMlCmd.eStateComplete) THEN
            _eState := E_DL_PackMlState.eStopped;
        END_IF

    E_DL_PackMlState.eAborting:                     // acting：急停执行（自动跃迁，无需 SC）
        _eState := E_DL_PackMlState.eAborted;

    E_DL_PackMlState.eAborted:                      // wait：已急停，仅 Clear/Reset 可退
        IF eCmd = E_DL_PackMlCmd.eClear THEN
            _eState := E_DL_PackMlState.eClearing;  // 恢复链第一步：清除去污
        ELSIF eCmd = E_DL_PackMlCmd.eReset THEN
            _eState := E_DL_PackMlState.eResetting;
        END_IF

    E_DL_PackMlState.eHolding:                      // acting：机内保持过渡
        IF bStateComplete OR (eCmd = E_DL_PackMlCmd.eStateComplete) THEN
            _eState := E_DL_PackMlState.eHeld;
        END_IF

    E_DL_PackMlState.eHeld:                         // wait：机内原因暂停
        IF eCmd = E_DL_PackMlCmd.eUnhold THEN
            _eState := E_DL_PackMlState.eUnholding;
        ELSIF eCmd = E_DL_PackMlCmd.eStop THEN
            _eState := E_DL_PackMlState.eStopping;
        ELSIF eCmd = E_DL_PackMlCmd.eAbort THEN
            _eState := E_DL_PackMlState.eAborting;
        END_IF

    E_DL_PackMlState.eUnholding:                    // acting：从保持回到执行
        IF bStateComplete OR (eCmd = E_DL_PackMlCmd.eStateComplete) THEN
            _eState := E_DL_PackMlState.eExecute;
        END_IF

    E_DL_PackMlState.eSuspending:                   // acting：机外暂停过渡
        IF bStateComplete OR (eCmd = E_DL_PackMlCmd.eStateComplete) THEN
            _eState := E_DL_PackMlState.eSuspended;
        END_IF

    E_DL_PackMlState.eUnsuspending:                 // acting：从挂起回到执行
        IF bStateComplete OR (eCmd = E_DL_PackMlCmd.eStateComplete) THEN
            _eState := E_DL_PackMlState.eExecute;
        END_IF

    E_DL_PackMlState.eResetting:                    // acting：复位子工序
        IF bStateComplete OR (eCmd = E_DL_PackMlCmd.eStateComplete) THEN
            _eState := E_DL_PackMlState.eIdle;      // Completed→Reset→Resetting→Idle 闭环
        END_IF

    E_DL_PackMlState.eCompleting:                   // acting：完工收尾子工序
        IF bStateComplete OR (eCmd = E_DL_PackMlCmd.eStateComplete) THEN
            _eState := E_DL_PackMlState.eCompleted;
        END_IF

    E_DL_PackMlState.eCompleted:                    // wait：批次完成
        IF eCmd = E_DL_PackMlCmd.eReset THEN
            _eState := E_DL_PackMlState.eResetting;
        ELSIF eCmd = E_DL_PackMlCmd.eClear THEN
            _eState := E_DL_PackMlState.eClearing;
        ELSIF eCmd = E_DL_PackMlCmd.eStop THEN
            _eState := E_DL_PackMlState.eStopping;
        ELSIF eCmd = E_DL_PackMlCmd.eAbort THEN
            _eState := E_DL_PackMlState.eAborting;
        END_IF

    ELSE
        // 非法状态兜底（故障级）：走 Aborting 路径
        _ePrevState := _eState;
        _eState := E_DL_PackMlState.eAborting;
        uErrorId := 16#0005_0201;

END_CASE

// 段 5｜跃迁刷新：仅真实跃迁时更新 ePrevState（Abort 复盘语义）
IF _eState <> _eStateOld THEN
    _ePrevState := _eStateOld;
END_IF

// 段 6｜状态出口映射：OEE 三位正交指示
eState := _eState;                                  // 当前状态出口
ePrevState := _ePrevState;                          // 前一状态出口
bInExecute := (_eState = E_DL_PackMlState.eExecute);              // Execute 计时位
bHeldByMachine := (_eState = E_DL_PackMlState.eHolding) OR (_eState = E_DL_PackMlState.eHeld)
                  OR (_eState = E_DL_PackMlState.eUnholding);     // 机内保持组
bSuspendedByLine := (_eState = E_DL_PackMlState.eSuspending) OR (_eState = E_DL_PackMlState.eSuspended)
                    OR (_eState = E_DL_PackMlState.eUnsuspending); // 机外挂起组
END_FUNCTION_BLOCK
